{attribute 'qualified_only'}
{attribute 'strict'}
TYPE E_Prod_Type :
(
	Marinade := 0,
	Color
);
END_TYPE

(* stored: Version 1.1.0.1, ProductVersion 3.1.4024.15
   DUT E_Prod_Type: Id {4b2219b2-a99b-4640-94be-15fe660a7a3c} *)
